(* IEC 61131-3 sources: 2026_Projet_YGO_ExcavatriceDragage/CODE_BACKUP/CODE_20260807_v0.5.25/DIAG, 5 files *)

(* ---- E_Diag_State.st ---- *)
(* ═══════════════════════════════════════════════════════════════
   🚦 E_Diag_State — Phases du cycle de diagnostic bus
   ═══════════════════════════════════════════════════════════════ *)
TYPE E_Diag_State :
(
    DISABLED   := 0,  (* Désactivé (surveillance non active) *)
    READY      := 1,  (* Opérationnel réel, pas de défaut *)
    INIT       := 2,  (* Initialisation / Recherche de réseau *)
    MONITORING := 3,  (* Surveillance active (états transitoires) *)
    ERROR      := 4,  (* Anomalie de communication *)
    SIMULATED  := 5   (* Bypass simulation ou bypass réseau IHM — pas le bus réel *)
);
END_TYPE

(* ---- ST_Diag_Device.st ---- *)
(* ═══════════════════════════════════════════════════════════════
   📡 ST_Diag_Device — Structure diagnostic d'un esclave ou bus
   ═══════════════════════════════════════════════════════════════ *)
TYPE ST_Diag_Device :
STRUCT
    Online         : BOOL;        (* Esclave visible sur le bus *)
    Operational    : BOOL;        (* Esclave en mode OP (opérationnel) *)
    Error          : BOOL;        (* Signal de défaut actif pour cet esclave *)
    ErrorId        : WORD;        (* Code défaut détaillé *)
    State          : E_Diag_State; (* Phase courante du cycle de diagnostic *)
    StateAtError   : E_Diag_State; (* Instantané de la phase lors de l'anomalie *)
END_STRUCT
END_TYPE

(* ---- FB_Diag_CanOpen.st ---- *)
(* ═══════════════════════════════════════════════════════════════
   📡 FB_Diag_CanOpen — Diagnostic bus CANopen / Joystick
   ───────────────────────────────────────────────────────────────
   📄 Docs : DOC/AF_Partie-02_Architecture_Programme_v3.1.md
              DOC/AF_Partie-06_Acquisition_Qualification_IO_v2.1.md §3
   🎯 Rôle : Décide Online/Operational et publie ST_Diag_Device.
      Distinction explicite dans State :
      - INIT       : pas encore online (ni réel, ni bypass)
      - SIMULATED  : bypass actif (simulation ou bypass réseau IHM)
      - READY      : bus réellement online
      - ERROR      : défaut détecté
   ═══════════════════════════════════════════════════════════════ *)
FUNCTION_BLOCK PUBLIC FB_Diag_CanOpen
VAR_INPUT
    Enable          : BOOL;        (* Active la surveillance CAN *)
    Reset           : BOOL;        (* Front d'acquittement des défauts *)
    CANbusStateRaw          : INT;          (* Valeur brute CANbus.GetBusState() (2 = ACTIVE) *)
    DeviceJoystickStateRaw  : DEVICE_STATE; (* Valeur brute JOY1.GetDeviceState() *)
    SimBypassActive         : BOOL;         (* TRUE = simulation active pour ce device *)
    NetworkBypassActive     : BOOL;         (* TRUE = bypass réseau global IHM *)
END_VAR
VAR_OUTPUT
    Ready           : BOOL;        (* Logique de surveillance active *)
    Busy            : BOOL;        (* Non utilisé (conformité interface) *)
    Done            : BOOL;        (* Non utilisé *)
    Error           : BOOL;        (* Présence anomalie de communication *)
    ErrorId         : WORD;        (* Code défaut global résumé *)
    State           : E_Diag_State; (* Phase courante (INIT/SIMULATED/READY/ERROR) *)
    StateAtError    : E_Diag_State; (* Phase figée à l'apparition de l'erreur *)
    DeviceCanOpenMaster : ST_Diag_Device;  (* Diagnostics bus CANopen *)
    DeviceJoystick  : ST_Diag_Device;  (* Diagnostics esclave Joystick *)
    (* Miroirs bruts lisibles directement sur l'instance *)
    CANbusStateRawOut         : INT;
    DeviceJoystickStateRawOut : DEVICE_STATE;
END_VAR
VAR
    ResetEdge       : R_TRIG;      (* Détecteur front de reset *)
    CANbusOnlineReal         : BOOL; (* Bus réellement actif, hors tout bypass *)
    DeviceJoystickOnlineReal : BOOL; (* Joystick réellement RUNNING, hors tout bypass *)
    BypassActive             : BOOL; (* Simulation OU bypass réseau IHM *)
    CANbusOnlineEff          : BOOL; (* Online effectif (réel OU bypass) *)
    DeviceJoystickOnlineEff  : BOOL; (* Operational effectif (réel OU bypass) *)
END_VAR

// 🛑 1. GATE : Désactivation logique si Enable = FALSE
IF NOT Enable THEN
    Ready := FALSE;
    State := E_Diag_State.DISABLED;
    DeviceJoystick.State := E_Diag_State.DISABLED;
    DeviceJoystick.Online := FALSE;
    DeviceJoystick.Operational := FALSE;
    DeviceJoystick.Error := FALSE;
    DeviceJoystick.ErrorId := 16#0000;
    DeviceCanOpenMaster.State := E_Diag_State.DISABLED;
    DeviceCanOpenMaster.Online := FALSE;
    DeviceCanOpenMaster.Operational := FALSE;
    Error := FALSE;
    ErrorId := 16#0000;
    CANbusStateRawOut := CANbusStateRaw;
    DeviceJoystickStateRawOut := DeviceJoystickStateRaw;
    RETURN;
END_IF;

Ready := TRUE;

// 🧮 2. INTERPRÉTATION DES VALEURS BRUTES
CANbusOnlineReal         := (CANbusStateRaw = 2);
DeviceJoystickOnlineReal := (DeviceJoystickStateRaw = DEVICE_STATE.RUNNING);
BypassActive             := SimBypassActive OR NetworkBypassActive;
CANbusOnlineEff          := CANbusOnlineReal OR BypassActive;
DeviceJoystickOnlineEff  := DeviceJoystickOnlineReal OR BypassActive;

// 🔑 3. RESET FRONT — Efface les défauts si la cause a disparu
ResetEdge(CLK := Reset);
IF ResetEdge.Q THEN
    IF (CANbusOnlineEff AND DeviceJoystickOnlineEff) THEN
        DeviceJoystick.ErrorId := 16#0000;
        StateAtError := E_Diag_State.DISABLED;
    END_IF;
END_IF;

// 🔍 4. DIAGNOSTIC JOYSTICK
// Bit 0 : Perte de communication CAN
IF NOT CANbusOnlineEff THEN
    DeviceJoystick.ErrorId := DeviceJoystick.ErrorId OR 16#0001;  (* Perte liaison CAN joystick *)
    DeviceJoystick.Online := FALSE;
ELSE
    DeviceJoystick.Online := TRUE;
    DeviceJoystick.ErrorId := DeviceJoystick.ErrorId AND 16#FFFE; (* Effacement auto si la liaison revient *)
END_IF;

// Bit 1 : Mode non-opérationnel (esclave CANopen en pré-op ou défaut)
IF NOT DeviceJoystickOnlineEff THEN
    DeviceJoystick.ErrorId := DeviceJoystick.ErrorId OR 16#0002;  (* Joystick pas opérationnel *)
    DeviceJoystick.Operational := FALSE;
ELSE
    DeviceJoystick.Operational := TRUE;
    DeviceJoystick.ErrorId := DeviceJoystick.ErrorId AND 16#FFFD; (* Effacement auto dès que RUNNING *)
END_IF;

// 🚦 5. MACHINE D'ÉTAT JOYSTICK
IF DeviceJoystick.ErrorId <> 0 THEN
    DeviceJoystick.State := E_Diag_State.ERROR;
    IF StateAtError = E_Diag_State.DISABLED THEN
        StateAtError := State;
    END_IF;
ELSIF NOT (DeviceJoystick.Online AND DeviceJoystick.Operational) THEN
    DeviceJoystick.State := E_Diag_State.INIT;
ELSIF BypassActive AND NOT (CANbusOnlineReal AND DeviceJoystickOnlineReal) THEN
    DeviceJoystick.State := E_Diag_State.SIMULATED;
ELSE
    DeviceJoystick.State := E_Diag_State.READY;
END_IF;

State := DeviceJoystick.State;

// 📤 6. SORTIES GLOBALES
DeviceJoystick.Error := (DeviceJoystick.ErrorId <> 0);
Error := DeviceJoystick.Error;
ErrorId := DeviceJoystick.ErrorId;

DeviceCanOpenMaster.Operational := CANbusOnlineEff;
DeviceCanOpenMaster.Online := CANbusOnlineEff;

IF NOT CANbusOnlineEff THEN
    DeviceCanOpenMaster.State := E_Diag_State.INIT;
ELSIF BypassActive AND NOT CANbusOnlineReal THEN
    DeviceCanOpenMaster.State := E_Diag_State.SIMULATED;
ELSE
    DeviceCanOpenMaster.State := E_Diag_State.READY;
END_IF;

// Miroirs bruts, toujours à jour
CANbusStateRawOut := CANbusStateRaw;
DeviceJoystickStateRawOut := DeviceJoystickStateRaw;

// Briques génériques pour conformité standard
Busy := FALSE;
Done := FALSE;

(* ---- FB_Diag_Ethercat.st ---- *)
(* ═══════════════════════════════════════════════════════════════
   📡 FB_Diag_Ethercat — Diagnostic bus EtherCAT (3 esclaves)
   ───────────────────────────────────────────────────────────────
   📄 Docs : DOC/AF_Partie-02_Architecture_Programme_v3.1.md
              DOC/AF_Partie-06_Acquisition_Qualification_IO_v2.1.md §3
   🎯 Rôle : Décide Online/Operational pour variateur M3 + codeurs M1/M2.
      Publie ST_Diag_Device par device + state global.
   ═══════════════════════════════════════════════════════════════ *)
FUNCTION_BLOCK PUBLIC FB_Diag_Ethercat
VAR_INPUT
    Enable              : BOOL;        (* Active la surveillance EtherCAT *)
    Reset               : BOOL;        (* Front d'acquittement des défauts *)

    (* Variateur M3 (AC600_ECAT_Drive) *)
    DeviceVariateurStateRaw     : DEVICE_STATE; (* Valeur brute AC600_ECAT_Drive.GetDeviceState() *)
    DeviceVariateurSimBypass    : BOOL;         (* TRUE = simulation active *)

    (* Encodeur M1 (COD1_CODEUR) *)
    DeviceEncoderM1StateRaw     : DEVICE_STATE; (* Valeur brute COD1_CODEUR.GetDeviceState() *)
    DeviceEncoderM1SimBypass    : BOOL;         (* TRUE = simulation active *)

    (* Encodeur M2 (COD2_CODEUR) *)
    DeviceEncoderM2StateRaw     : DEVICE_STATE; (* Valeur brute COD2_CODEUR.GetDeviceState() *)
    DeviceEncoderM2SimBypass    : BOOL;         (* TRUE = simulation active *)

    NetworkBypassActive         : BOOL;         (* TRUE = bypass réseau global IHM *)
END_VAR
VAR_OUTPUT
    Ready               : BOOL;        (* Logique de surveillance active *)
    Busy                : BOOL;        (* Non utilisé (conformité) *)
    Done                : BOOL;        (* Non utilisé *)
    Error               : BOOL;        (* Résumé anomalie de communication bus *)
    ErrorId             : WORD;        (* Code défaut global résumé *)
    State               : E_Diag_State; (* Phase courante du diagnostic global — voir en-tête *)
    StateAtError        : E_Diag_State; (* Phase figée à l'apparition de l'erreur *)
    DeviceEthercatMaster : ST_Diag_Device; (* Diagnostics bus EtherCAT *)
    DeviceVariateur     : ST_Diag_Device;  (* Diagnostics esclave AC600 *)
    DeviceEncoderM1     : ST_Diag_Device;  (* Diagnostics esclave COD1 *)
    DeviceEncoderM2     : ST_Diag_Device;  (* Diagnostics esclave COD2 *)
    (* Miroirs bruts lisibles directement sur l'instance *)
    DeviceVariateurStateRawOut : DEVICE_STATE;
    DeviceEncoderM1StateRawOut : DEVICE_STATE;
    DeviceEncoderM2StateRawOut : DEVICE_STATE;
END_VAR
VAR
    ResetEdge           : R_TRIG;      (* Détecteur front de reset *)
    VariateurOnlineReal  : BOOL; (* GetDeviceState() = RUNNING, hors tout bypass *)
    EncoderM1OnlineReal  : BOOL;
    EncoderM2OnlineReal  : BOOL;
    VariateurBypass      : BOOL; (* Simulation OU bypass réseau IHM, pour ce device *)
    EncoderM1Bypass      : BOOL;
    EncoderM2Bypass      : BOOL;
    VariateurOnlineEff   : BOOL; (* Online effectif (réel OU bypass) *)
    EncoderM1OnlineEff   : BOOL;
    EncoderM2OnlineEff   : BOOL;
END_VAR

// 🛑 1. GATE : Désactivation si Enable = FALSE
IF NOT Enable THEN
    Ready := FALSE;
    State := E_Diag_State.DISABLED;
    DeviceVariateur.State := E_Diag_State.DISABLED;
    DeviceEncoderM1.State := E_Diag_State.DISABLED;
    DeviceEncoderM2.State := E_Diag_State.DISABLED;
    DeviceVariateur.Online := FALSE;
    DeviceEncoderM1.Online := FALSE;
    DeviceEncoderM2.Online := FALSE;
    DeviceVariateur.Operational := FALSE;
    DeviceEncoderM1.Operational := FALSE;
    DeviceEncoderM2.Operational := FALSE;
    DeviceVariateur.Error := FALSE;
    DeviceEncoderM1.Error := FALSE;
    DeviceEncoderM2.Error := FALSE;
    Error := FALSE;
    ErrorId := 16#0000;
    DeviceEthercatMaster.State := E_Diag_State.DISABLED;
    DeviceEthercatMaster.Online := FALSE;
    DeviceEthercatMaster.Operational := FALSE;
    DeviceVariateurStateRawOut := DeviceVariateurStateRaw;
    DeviceEncoderM1StateRawOut := DeviceEncoderM1StateRaw;
    DeviceEncoderM2StateRawOut := DeviceEncoderM2StateRaw;
    RETURN;
END_IF;

Ready := TRUE;

// 🧮 2. INTERPRÉTATION DES VALEURS BRUTES
VariateurOnlineReal := (DeviceVariateurStateRaw = DEVICE_STATE.RUNNING);
EncoderM1OnlineReal := (DeviceEncoderM1StateRaw = DEVICE_STATE.RUNNING);
EncoderM2OnlineReal := (DeviceEncoderM2StateRaw = DEVICE_STATE.RUNNING);

VariateurBypass := DeviceVariateurSimBypass OR NetworkBypassActive;
EncoderM1Bypass := DeviceEncoderM1SimBypass OR NetworkBypassActive;
EncoderM2Bypass := DeviceEncoderM2SimBypass OR NetworkBypassActive;

VariateurOnlineEff := VariateurOnlineReal OR VariateurBypass;
EncoderM1OnlineEff := EncoderM1OnlineReal OR EncoderM1Bypass;
EncoderM2OnlineEff := EncoderM2OnlineReal OR EncoderM2Bypass;

// 🔑 3. RESET FRONT
ResetEdge(CLK := Reset);

// 🔍 4. DIAGNOSTIC VARIATEUR (AC600_ECAT_Drive / Translation M3)
DeviceVariateur.Online := VariateurOnlineEff;
DeviceVariateur.Operational := VariateurOnlineEff;

IF NOT DeviceVariateur.Online THEN
    DeviceVariateur.ErrorId := DeviceVariateur.ErrorId OR 16#0010;  (* Perte liaison physique variateur *)
ELSE
    DeviceVariateur.ErrorId := DeviceVariateur.ErrorId AND 16#FFEF; (* Effacement auto dès que RUNNING *)
END_IF;

// 🔍 5. DIAGNOSTIC ENCODEUR M1 (COD1_CODEUR / WinchM1)
DeviceEncoderM1.Online := EncoderM1OnlineEff;
DeviceEncoderM1.Operational := EncoderM1OnlineEff;

IF NOT DeviceEncoderM1.Online THEN
    DeviceEncoderM1.ErrorId := DeviceEncoderM1.ErrorId OR 16#0020;  (* Perte liaison encodeur M1 *)
ELSE
    DeviceEncoderM1.ErrorId := DeviceEncoderM1.ErrorId AND 16#FFDF; (* Effacement auto dès que RUNNING *)
END_IF;

// 🔍 6. DIAGNOSTIC ENCODEUR M2 (COD2_CODEUR / WinchM2)
DeviceEncoderM2.Online := EncoderM2OnlineEff;
DeviceEncoderM2.Operational := EncoderM2OnlineEff;

IF NOT DeviceEncoderM2.Online THEN
    DeviceEncoderM2.ErrorId := DeviceEncoderM2.ErrorId OR 16#0030;  (* Perte liaison encodeur M2 *)
ELSE
    DeviceEncoderM2.ErrorId := DeviceEncoderM2.ErrorId AND 16#FFCF; (* Effacement auto dès que RUNNING *)
END_IF;

// 🚦 7. STATE MACHINES DE CHAQUE APPAREIL
IF DeviceVariateur.ErrorId <> 0 THEN
    DeviceVariateur.State := E_Diag_State.ERROR;
ELSIF NOT VariateurOnlineEff THEN
    DeviceVariateur.State := E_Diag_State.INIT;
ELSIF VariateurBypass AND NOT VariateurOnlineReal THEN
    DeviceVariateur.State := E_Diag_State.SIMULATED;
ELSE
    DeviceVariateur.State := E_Diag_State.READY;
END_IF;

IF DeviceEncoderM1.ErrorId <> 0 THEN
    DeviceEncoderM1.State := E_Diag_State.ERROR;
ELSIF NOT EncoderM1OnlineEff THEN
    DeviceEncoderM1.State := E_Diag_State.INIT;
ELSIF EncoderM1Bypass AND NOT EncoderM1OnlineReal THEN
    DeviceEncoderM1.State := E_Diag_State.SIMULATED;
ELSE
    DeviceEncoderM1.State := E_Diag_State.READY;
END_IF;

IF DeviceEncoderM2.ErrorId <> 0 THEN
    DeviceEncoderM2.State := E_Diag_State.ERROR;
ELSIF NOT EncoderM2OnlineEff THEN
    DeviceEncoderM2.State := E_Diag_State.INIT;
ELSIF EncoderM2Bypass AND NOT EncoderM2OnlineReal THEN
    DeviceEncoderM2.State := E_Diag_State.SIMULATED;
ELSE
    DeviceEncoderM2.State := E_Diag_State.READY;
END_IF;

// Fige la phase du diagnostic global sur le premier défaut
IF (DeviceVariateur.ErrorId <> 0 OR DeviceEncoderM1.ErrorId <> 0 OR DeviceEncoderM2.ErrorId <> 0) THEN
    IF StateAtError = E_Diag_State.DISABLED THEN
        StateAtError := State;
    END_IF;
END_IF;

// 📤 8. RÉSUMÉ ET DÉFAUTS
DeviceVariateur.Error := (DeviceVariateur.ErrorId <> 0);
DeviceEncoderM1.Error := (DeviceEncoderM1.ErrorId <> 0);
DeviceEncoderM2.Error := (DeviceEncoderM2.ErrorId <> 0);

Error := (DeviceVariateur.Error OR DeviceEncoderM1.Error OR DeviceEncoderM2.Error);

ErrorId := 16#0000;
IF DeviceVariateur.Error THEN
    ErrorId := ErrorId OR 16#00F0;
END_IF;
IF DeviceEncoderM1.Error THEN
    ErrorId := ErrorId OR 16#0F00;
END_IF;
IF DeviceEncoderM2.Error THEN
    ErrorId := ErrorId OR 16#F000;
END_IF;

IF Error THEN
    State := E_Diag_State.ERROR;
ELSIF NOT (VariateurOnlineEff AND EncoderM1OnlineEff AND EncoderM2OnlineEff) THEN
    State := E_Diag_State.INIT;
ELSIF (VariateurBypass OR EncoderM1Bypass OR EncoderM2Bypass)
      AND NOT (VariateurOnlineReal AND EncoderM1OnlineReal AND EncoderM2OnlineReal) THEN
    State := E_Diag_State.SIMULATED;
ELSE
    State := E_Diag_State.READY;
END_IF;

DeviceEthercatMaster.Online := VariateurOnlineEff AND EncoderM1OnlineEff AND EncoderM2OnlineEff;
DeviceEthercatMaster.Operational := DeviceEthercatMaster.Online;

DeviceVariateurStateRawOut := DeviceVariateurStateRaw;
DeviceEncoderM1StateRawOut := DeviceEncoderM1StateRaw;
DeviceEncoderM2StateRawOut := DeviceEncoderM2StateRaw;

Busy := FALSE;
Done := FALSE;

(* ---- FB_Diag_IhmHeartbeat.st ---- *)
(* ═══════════════════════════════════════════════════════════════
   💓 FB_Diag_IhmHeartbeat — Surveillance bidirectionnelle IHM↔PLC
   ───────────────────────────────────────────────────────────────
   📄 Doc : DOC/AF_Partie-07_Interface_IHM_v2.0.md (mise à jour Heartbeat requise)
   🧩 Brique réduite : surveille le toggle IHM, génère le toggle PLC
      et expose un diagnostic. Ne produit ni SafeStop ni PowerCutOff.
   🛡️ Les FB_Safety_Winch / FB_Safety_Translation restent propriétaires
      de leurs réactions métier.
   ═══════════════════════════════════════════════════════════════ *)

FUNCTION_BLOCK PUBLIC FB_Diag_IhmHeartbeat
VAR_INPUT
    Enable              : BOOL;              // Active la surveillance ; FALSE = IHM non valide
    TglHeartbeatIhm  : BOOL;              // Toggle IHM, inversion attendue toutes les 500 ms
    IhmTimeout          : TIME := T#2s;     // Absence maximale de front IHM
    PlcTogglePeriod     : TIME := T#500ms;  // Période du clignotant PLC
END_VAR
VAR_OUTPUT
    HeartbeatIhmOk      : BOOL;              // TRUE après front IHM post-boot et avant timeout
    HeartbeatIhmTimeout : BOOL;              // TRUE = aucun front IHM depuis IhmTimeout
    TglHeartbeatPlc  : BOOL;              // Clignotant PLC à superviser côté IHM
    TimeSinceIhmEdge    : TIME;              // Diagnostic : temps depuis le dernier front IHM
END_VAR
VAR
    LastIhmToggle       : BOOL;
    IhmEdgeSeen         : BOOL;              // Interdit de valider une valeur RETAIN au boot
    IhmEdgeDetected     : BOOL;
    IhmTimeoutTon       : TON;
    PlcToggleTon        : TON;
END_VAR

// === IMPLEMENTATION ===

// 🛑 Sans Enable, aucune valeur mémorisée ne peut déclarer l'IHM valide.
IF NOT Enable THEN
    HeartbeatIhmOk := FALSE;
    HeartbeatIhmTimeout := TRUE;
    TglHeartbeatPlc := FALSE;
    TimeSinceIhmEdge := T#0s;
    LastIhmToggle := TglHeartbeatIhm;
    IhmEdgeSeen := FALSE;
    IhmTimeoutTon(IN := FALSE, PT := IhmTimeout);
    PlcToggleTon(IN := FALSE, PT := PlcTogglePeriod);
    RETURN;
END_IF;

// 📥 Front par comparaison : l'IHM écrit un BOOL toggle, pas une impulsion courte.
IhmEdgeDetected := (TglHeartbeatIhm <> LastIhmToggle);
LastIhmToggle := TglHeartbeatIhm;
IF IhmEdgeDetected THEN
    IhmEdgeSeen := TRUE;
END_IF;

// ⏱️ Le timer repart à chaque front. Au boot, il atteint le timeout au bout de IhmTimeout.
// HeartbeatIhmOk reste TRUE tant que le timeout n'est pas expiré (boot propre sans alarme au scan 1).
IhmTimeoutTon(IN := NOT IhmEdgeDetected, PT := IhmTimeout);
TimeSinceIhmEdge := IhmTimeoutTon.ET;
HeartbeatIhmTimeout := IhmTimeoutTon.Q;
HeartbeatIhmOk := NOT HeartbeatIhmTimeout;

// 💡 Clignotant PLC indépendant : information de vie pour l'IHM, jamais signal Safety autonome.
PlcToggleTon(IN := NOT PlcToggleTon.Q, PT := PlcTogglePeriod);
IF PlcToggleTon.Q THEN
    TglHeartbeatPlc := NOT TglHeartbeatPlc;
END_IF;
